(* IEC 61131-3 sources: JingjiangMoonbox/Application/Application/任务列表/Main_Task/GNS_MAP, 4 files *)

(* ---- KS_CreatGantryAxisInf.st ---- *)
(*@CES
Name=KS_CreatGantryAxisInf
Type=FunctionBlock
TypeGuid=6f9dac99-8de1-4efc-8465-68ac443b7d08
Guid=f41a9b20-4237-42b7-ab68-52a2ca659d0d
HasDeclaration=True
HasImplementation=True
*)
{DECLARATION}
FUNCTION KS_CreatGantryAxisInf : BOOL
(*获取龙门轴信息*)
VAR_INPUT
	(*输入*)
	i_pstStSysStationInf 	: POINTER TO StSysStationInf;
	(*输出*)
	i_pstStSysGantryAxisInf : POINTER TO StSysGantryAxisInf;
END_VAR
VAR
	in					: INT;
	pstStStationInf		: POINTER TO StStationInf;
	pstStGantryAxisInf	: POINTER TO StGantryAxisInf;
	(*龙门轴信息地址@索引为轴id,最大15*)
	(*每个轴2个龙门@二维数组里的1是版辊、2是网纹辊*)
	apstStGantryAxisInf	: ARRAY [1..20,1..2] OF POINTER TO StGantryAxisInf:=[40(0)];
	iGantryAxisNum		: INT := 0;(*龙门轴个数*)
	iMaxGantryAxisNum	: INT;
	iLogicAxisId		: INT;(*逻辑轴id*)
	iLogicAxisIdSuperPos: INT;(*叠加轴id*)
	iMoveType			: stEnumMoveType;(*运动类型*)
	iAxisId				: stEnumAxisId;
	iStaitonFuncId		: stEnumFuncId;
	iCoreId				: INT;
	iIndexTmp			: INT;(*数组索引*)
END_VAR
{IMPLEMENTATION}
IF i_pstStSysStationInf<>0 AND i_pstStSysGantryAxisInf<>0 THEN
	(*龙门组个数*)
	iMaxGantryAxisNum:=SIZEOF(i_pstStSysGantryAxisInf^.astGantryAxisInf)/SIZEOF(i_pstStSysGantryAxisInf^.astGantryAxisInf[1]);
	(*初始化*)
	FOR iN:=1 TO iMaxGantryAxisNum BY 1 DO
		KS_InitGantryAxisInf(ADR(i_pstStSysGantryAxisInf^.astGantryAxisInf[iN]));
	END_FOR
	(*从系统架构中找龙门轴*)
	FOR in:=1 TO i_pstStSysStationInf^.byStationNum BY 1 DO
		pstStStationInf:=ADR(i_pstStSysStationInf^.astStationInf[iN]);
		IF pstStStationInf^.xValid THEN
			iAxisId					:=pstStStationInf^.iAxisId;
			iLogicAxisId			:=pstStStationInf^.iLogicAxisId;
			iLogicAxisIdSuperPos	:=pstStStationInf^.iLogicAxisIdSuperPos;
			iMoveType				:=pstStStationInf^.iMoveType;
			iStaitonFuncId			:=pstStStationInf^.iFuncId;
			iCoreId					:=pstStStationInf^.iCoreId_LogicAxis;
			IF KS_IsUnitAxisId(iAxisId)THEN(*是色组*)
				IF iMoveType = MOVETYPE_GANTRY THEN(*龙门轴*)
					IF iStaitonFuncId = FUNCID_PRNROLLER_PRESSURE_M OR
						iStaitonFuncId = FUNCID_PRNROLLER_PRESSURE_G THEN(*印刷辊龙门*)
						iIndexTmp:=1;
					ELSE(*else都认为是网纹辊龙门*)
						iIndexTmp:=2;
					END_IF

					IF apstStGantryAxisInf[iAxisId,iIndexTmp] = 0 THEN
						iGantryAxisNum:=iGantryAxisNum+1;
						(*获取龙门轴需要的信息*)
						(*写入的结构体地址获取*)
						IF iGantryAxisNum<=iMaxGantryAxisNum THEN
							pstStGantryAxisInf:=ADR(i_pstStSysGantryAxisInf^.astGantryAxisInf[iGantryAxisNum]);
						ELSE(*超限了|退出*)
							EXIT;
						END_IF
						apstStGantryAxisInf[iAxisId,iIndexTmp]:=ADR(i_pstStSysGantryAxisInf^.astGantryAxisInf[iGantryAxisNum]);
					END_IF

					(*获取地址*)
					pstStGantryAxisInf:=apstStGantryAxisInf[iAxisId,iIndexTmp];
					IF pstStGantryAxisInf<>0 THEN(*地址合法*)
						pstStGantryAxisInf^.iAxisId:=iAxisId;
						pstStGantryAxisInf^.iCoreId:=iCoreId;(*龙门站必须是一个核|所以不用区分*)

						CASE iStaitonFuncId OF
							FUNCID_PRNROLLER_PRESSURE_M:(*版辊压力|操作侧@叠加轴id在m侧的数据里*)
								pstStGantryAxisInf^.iFuncId					:=FUNCID_PRNROLLER_GANTRY;
								pstStGantryAxisInf^.iLogicAxisId_M			:=iLogicAxisId;
								pstStGantryAxisInf^.iLogicAxisId_SuperPos	:=iLogicAxisIdSuperPos;
							FUNCID_PRNROLLER_PRESSURE_G:
								pstStGantryAxisInf^.iFuncId					:=FUNCID_PRNROLLER_GANTRY;
								pstStGantryAxisInf^.iLogicAxisId_G			:=pstStStationInf^.iLogicAxisId;
							FUNCID_NETROLLER_PRESSURE_M:(*网辊压力|操作侧@叠加轴id在m侧的数据里*)
								pstStGantryAxisInf^.iFuncId					:=FUNCID_NETROLLER_GANTRY;
								pstStGantryAxisInf^.iLogicAxisId_M			:=iLogicAxisId;
								pstStGantryAxisInf^.iLogicAxisId_SuperPos	:=iLogicAxisIdSuperPos;
							FUNCID_NETROLLER_PRESSURE_G:
								pstStGantryAxisInf^.iFuncId					:=FUNCID_NETROLLER_GANTRY;
								pstStGantryAxisInf^.iLogicAxisId_G			:=pstStStationInf^.iLogicAxisId;
						ELSE;(*不是压力的就不理会了*)
						END_CASE
					END_IF
				ELSE(*不是龙门轴不理会*);
				END_IF
			END_IF(*不是色组就不理会了*);
		END_IF
	END_FOR
	i_pstStSysGantryAxisInf^.byGantryAxisNum:=INT_TO_BYTE(iGantryAxisNum);

	(*非法值检测*)
	FOR iN:=1 TO iGantryAxisNum BY 1 DO
		pstStGantryAxisInf:=ADR(i_pstStSysGantryAxisInf^.astGantryAxisInf[iN]);
		pstStGantryAxisInf^.xValid:=TRUE;
		IF pstStGantryAxisInf^.iAxisId=-1 OR
			pstStGantryAxisInf^.iCoreId=-1 OR
			pstStGantryAxisInf^.iFuncId=FUNCID_NULL OR
			pstStGantryAxisInf^.iLogicAxisId_G=-1 OR
			pstStGantryAxisInf^.iLogicAxisId_M=-1 OR
			pstStGantryAxisInf^.iLogicAxisId_SuperPos=-1 THEN
			pstStGantryAxisInf^.xValid:=FALSE;
		END_IF
	END_FOR
END_IF

(* ---- KS_CreatMap.st ---- *)
(*@CES
Name=KS_CreatMap
Type=FunctionBlock
TypeGuid=6f9dac99-8de1-4efc-8465-68ac443b7d08
Guid=61e29dc5-e287-4a1a-b094-66cbd5c76957
HasDeclaration=True
HasImplementation=True
*)
{DECLARATION}
FUNCTION KS_CreatMap : BOOL
(*创建映射表@触发执行|初始化获取到了站列表后执行一次就行*)
(*对应关系参考站号定义、xml分配文件*)
(*新的架构需要同步修改KS_CreatStationIdMap\KS_GetLogicAxisInfByStationIdForMap*)
(*2026.5.20.140844 by liu.yt 调整接口为系统列表结构体*)
VAR_INPUT
	i_xEn					: BOOL;(*创建使能@事件触发*)
	i_xUseRealStation		: BOOL;(*使用实际站创建*)
	(*根据系统架构创建*)
	i_iMachineryType		: stEuumMachineryType;(*机器类型*)
(*
	i_xIsDualUwRw			: BOOL;(*双收双放机型|*)
	i_xIfOfIsGlink			: BOOL;(*收放牵是glink站*)
	i_xUwRwIsGlink			: BOOL;(*收放料是glink站*)
	i_xPrnPressureIsGlink	: BOOL;(*印刷辊的压力辊是glink站*)
	i_xNetPressureIsGlink	: BOOL;(*网纹辊的压力辊是glink站*)
*)

	(*系统中实际站信息*)
	i_byStationIdNum		: BYTE;(*站的个数*)
	//i_piStationIdList		: POINTER TO INT;(*站id列表*)
	i_pstStStationInfo_KS	: POINTER TO StStationInfo_KS;(*固高函数获取的系统站信息@2026.5.20.140838 by liu.yt*)
	(*输出列表*)
	i_pstStSysStationInf	: POINTER TO StSysStationInf;
END_VAR
VAR
	iN					: INT;
	iAxisId				: stEnumAxisId;
	piTmp				: POINTER TO INT;
	pwTmp				: POINTER TO WORD;
	iStationInflenth	: INT;
	iStationNum			: INT;(*站的个数*)
	iValidStationNum	: INT;(*有效站个数*)
	aiStationidList		: ARRAY [1..256] OF INT;
	wStationType		: WORD;(*站的类型*)
	awStationType		: ARRAY [1..256] OF WORD;(*2026.5.20.141316 by liu.yt*)
	pstStationInf		: POINTER TO StStationInf;
	iFuncId				: stEnumFuncId;(*只针对色组轴*)
	iMoveType			: stEnumMoveType;(*运动的类型也可以获取*)
	iStationId			: INT;
	iCoreId				: INT:=-1;
	iLogicAxisIdSuperPos: INT:=-1;
	iLogicAxisId		: INT:=-1;
	(*不同的机型必须要显式赋值*)
	(*色组数@默认写的是机组式柔印+4压力电机*)
	iUnitNum			: INT:=10;
	iMachineryType		: stEuumMachineryType;
END_VAR
{IMPLEMENTATION}
IF i_xEn THEN
	iStationInflenth:=SIZEOF(i_pstStSysStationInf^.astStationInf) /
						SIZEOF(i_pstStSysStationInf^.astStationInf[1]);
	iMachineryType:=i_iMachineryType;
	(*获取站列表和个数*)
	IF i_xUseRealStation THEN
		(*2026.5.20.141002 by liu.yt*)
		//iStationNum:=BYTE_TO_INT(i_byStationIdNum);
		(*piTmp:=i_piStationIdList;*)
		iStationNum:=i_pstStStationInfo_KS^.iStationNum;
		piTmp:=ADR(i_pstStStationInfo_KS^.aiStationId_List);
		pwTmp:=ADR(i_pstStStationInfo_KS^.awStation_Type);
		FOR iN:=1 TO iStationNum BY 1 DO
			(*列表获取@2026.5.20.141347 by liu.yt*)
			aiStationidList[iN]:=piTmp^;
			piTmp:=piTmp+SIZEOF(piTmp^);
			(*站类型获取@2026.5.20.141359 by liu.yt*)
			awStationType[iN]:=pwTmp^;
			pwTmp:=pwTmp+SIZEOF(pwTmp^);
		END_FOR
	ELSE
		iStationNum:=255(*iStationInflenth*);
		IF iStationNum<=255 THEN
			FOR iN:=1 TO iStationNum BY 1 DO
				aiStationidList[iN]:=iN;
			END_FOR
		END_IF
	END_IF
	(*初始化@结构体数据*)
	i_pstStSysStationInf^.byStationNum:=0;
	FOR iN:=1 TO iStationInflenth BY 1 DO
		pstStationInf:=ADR(i_pstStSysStationInf^.astStationInf[iN]);
		KS_InitStationInf(pstStationInf);
	END_FOR

	iValidStationNum:=0;
(*	IF NOT i_xIsDualUwRw THEN(*常规机型*)*)
		(*按照*)
		CASE iMachineryType OF
			MACHINERYTYPE_ROTOGRAVE:(*凹印机*);
			MACHINERYTYPE_FELXO_INLINE,(*机组式柔印*)
			MACHINERYTYPE_FELXO_INLINE_ONEBOTOMROLLER:(*机组式柔印@单底辊*)
				(*按照10色，带龙门压力，横向配置@压力轴的个数限制了最大色组数只能为10个*)
				iUnitNum:=10;(*4电机压力限制最大只能10色*)
				(*处理map*)
				FOR iN:=1 TO iStationNum BY 1 DO
					iStationId:=aiStationidList[iN];
					wStationType:=awStationType[iN];
					(*获取轴信息*)
					iAxisId:=KS_GetAxisInfByStationIdForMap(iStationId,ADR(iFuncId),ADR(iMoveType));
					(*站号在表里,就输出有效标志*)
					IF iAxisId<>AXISID_INVALID THEN
						IF iAxisId > iUnitNum AND iAxisId <= AXISID_15U THEN(*非法轴id就剔除*);
						ELSE;
							iValidStationNum:=iValidStationNum+1;
							IF iValidStationNum<=iStationInflenth THEN
								pstStationInf:=ADR(i_pstStSysStationInf^.astStationInf[iValidStationNum]);
								pstStationInf^.xValid:=TRUE;
								pstStationInf^.iAxisId:=iAxisId;
								pstStationInf^.iStationId:=iStationId;
								pstStationInf^.iFuncId:=iFuncId;
								pstStationInf^.iMoveType:=iMoveType;
								pstStationInf^.udiStationType:=WORD_TO_UDINT(wStationType);(*2026.5.20.161045 by liu.yt*)
								(*运控信息获取*)
								iLogicAxisId:=
									KS_GetLogicAxisInfByStationIdForMap(
												iStationId(*i_iStationId*),
												iMachineryType(*i_iMachineryType*),
												ADR(iCoreId)(*i_piCoreId*),
												ADR(iLogicAxisIdSuperPos)(*i_piLogicAxisIdSuperPos*));

								pstStationInf^.iCoreId_LogicAxis			:=iCoreId;
								pstStationInf^.iCoreId_LogicAxisSuperPos	:=iCoreId;
								pstStationInf^.iLogicAxisId					:=iLogicAxisId;
								pstStationInf^.iLogicAxisIdSuperPos			:=iLogicAxisIdSuperPos;
							ELSE;(*超过最大索引了*)
								iValidStationNum:=iStationInflenth;(*站个数最大就是数组长度*)
							END_IF
						END_IF
					END_IF
				END_FOR

			MACHINERYTYPE_FELXO_CL:(*卫星式柔印*);
			MACHINERYTYPE_OFFSET:(*胶印机*);
		ELSE;
		END_CASE
(*
	ELSE;
	END_IF
*)
	i_pstStSysStationInf^.byStationNum:=INT_TO_BYTE(iValidStationNum);
END_IF

//2025.12.27.142131 | + 机器类型搞个变量单独弄出来
g_iMachineryType := i_iMachineryType;

(* ---- KS_GetAxisIdForMotByStation_Gantry.st ---- *)
(*@CES
Name=KS_GetAxisIdForMotByStation_Gantry
Type=FunctionBlock
TypeGuid=6f9dac99-8de1-4efc-8465-68ac443b7d08
Guid=cde7d95e-737e-4f32-881d-821472d364d1
HasDeclaration=True
HasImplementation=True
*)
{DECLARATION}
FUNCTION KS_GetAxisIdForMotByStation_Gantry : BOOL
(*转换为火眼原来设计的数据项，并输出。方便程序移植*)
VAR_INPUT
	i_iStationId			: INT;
	i_piAxisId				: POINTER TO INT;(*逻辑轴id*)
	i_piTypeId				: POINTER TO ENUM_AXISTYPE;(*类型id*)
	i_piUnitId				: POINTER TO INT;(*色组id*)
	i_piCoreId				: POINTER TO INT;(*核id*)
	i_piGroupId			 	: POINTER TO INT;(*组id*)
	i_piAdjAxisId			: POINTER TO INT;(*调整轴id*)
	(*系统列表*)
	i_pstStSysStationInf	: POINTER TO StSysStationInf;
	i_pstStSysGantryAxisInf	: POINTER TO StSysGantryAxisInf;
END_VAR
VAR
	iN					:  INT;
	xResult				:  BOOL:=FALSE;
	iAxisId				:  INT:=-1;(*逻辑轴id*)
	iTypeId				:  ENUM_AXISTYPE:=TYPE_NULL;(*类型id*)
	iUnitId				:  INT:=-1;(*色组id*)
	iCoreId				:  INT:=-1;(*核id*)
	iGroupId			:  INT:=-1;(*组id*)
	iAdjAxisId			:  INT:=-1;(*调整轴id*)
	pstStStationInf 	:  POINTER TO StStationInf;
	pstStGantryAxisInf	:  POINTER TO StGantryAxisInf;
END_VAR

{IMPLEMENTATION}
IF i_pstStSysStationInf <>0 AND i_pstStSysGantryAxisInf <> 0 THEN
	IF i_iStationId>0 AND i_iStationId<255 THEN(*站号合法性判断*)
		FOR iN:=1 TO i_pstStSysStationInf^.byStationNum BY 1 DO
			pstStStationInf:=ADR(i_pstStSysStationInf^.astStationInf[iN]);
			IF pstStStationInf^.xValid THEN
				IF i_iStationId = pstStStationInf^.iStationId THEN(*找到了*)
					xResult:=TRUE;
					iAxisId:=pstStStationInf^.iLogicAxisId;(*逻辑轴id*)
					IF KS_IsUnitAxisId(pstStStationInf^.iAxisId) THEN(*检查是不是色组的枚举*)
						iUnitId:=pstStStationInf^.iAxisId;
					END_IF
					iCoreId:=pstStStationInf^.iCoreId_LogicAxis;(*核id*)
					iAdjAxisId:=pstStStationInf^.iLogicAxisIdSuperPos;(*叠加轴id*)
					EXIT;
				END_IF
			END_IF
		END_FOR
	END_IF

	(*type处理*)
	iTypeId:=TYPE_NULL;
	IF xResult THEN
		CASE pstStStationInf^.iAxisId OF
			AXISID_UWA:		iTypeId:=TYPE_UNWIND_A_I;
			AXISID_UWB:		iTypeId:=TYPE_UNWIND_B_I;
			AXISID_RWA:		iTypeId:=TYPE_REWIND_A_I;
			AXISID_RWB:		iTypeId:=TYPE_REWIND_B_I;
			AXISID_IF:		iTypeId:=TYPE_INFEED_I;
			AXISID_OF:		iTypeId:=TYPE_OUTFEED_I;
			AXISID_UWA_II:	iTypeId:=TYPE_UNWIND_A_II;
			AXISID_UWB_II:	iTypeId:=TYPE_UNWIND_B_II;
			AXISID_RWA_II:	iTypeId:=TYPE_REWIND_A_II;
			AXISID_RWB_II:	iTypeId:=TYPE_REWIND_B_II;
			AXISID_IF_II:	iTypeId:=TYPE_INFEED_II;
			AXISID_OF_II:	iTypeId:=TYPE_OUTFEED_II;
			AXISID_CENTER:  iTypeId:=TYPE_CENTRAL_I;(*只处理单系中心辊*)
		ELSE
			(*色组*)
			IF  KS_IsUnitAxisId(pstStStationInf^.iAxisId) THEN
				CASE pstStStationInf^.iFuncId OF
					FUNCID_PRNROLLER: 				iTypeId:=TYPE_UNIT_PRN;
					FUNCID_NETROLLER: 				iTypeId:=TYPE_UNIT_NET;
					FUNCID_BOTTOMROLLER: 			iTypeId:=TYPE_UNIT_BOTTOM;
					FUNCID_PRNROLLER_PRESSURE_M: 	iTypeId:=TYPE_UNIT_PRN_PRESS_MASTER;
					FUNCID_PRNROLLER_PRESSURE_G: 	iTypeId:=TYPE_UNIT_PRN_PRESS_G;
					FUNCID_NETROLLER_PRESSURE_M: 	iTypeId:=TYPE_UNIT_NET_PRESS_MASTER;
					FUNCID_NETROLLER_PRESSURE_G: 	iTypeId:=TYPE_UNIT_NET_PRESS_G;
					FUNCID_HORZ: 					iTypeId:=TYPE_UNIT_HORIZ;
				ELSE;
				END_CASE
			END_IF
		END_CASE
	END_IF

	//龙门处理
	FOR iN:=1 TO i_pstStSysGantryAxisInf^.byGantryAxisNum BY 1 DO
		pstStGantryAxisInf := ADR(i_pstStSysGantryAxisInf^.astGantryAxisInf[iN]);
		IF  pstStGantryAxisInf^.xValid THEN
			IF iUnitId = pstStGantryAxisInf^.iAxisId THEN
				IF pstStGantryAxisInf^.iFuncId = FUNCID_PRNROLLER_GANTRY THEN
					IF iTypeId = TYPE_UNIT_PRN_PRESS_MASTER OR iTypeId = TYPE_UNIT_PRN_PRESS_G THEN
						iGroupId := iN;
						EXIT;
					END_IF
				ELSIF pstStGantryAxisInf^.iFuncId = FUNCID_NETROLLER_GANTRY THEN
					IF iTypeId = TYPE_UNIT_NET_PRESS_MASTER OR iTypeId = TYPE_UNIT_NET_PRESS_G THEN
						iGroupId := iN;
						EXIT;
					END_IF
				END_IF
			END_IF
		END_IF
	END_FOR
END_IF

IF i_piAxisId<>0 THEN
	i_piAxisId^:=iAxisId;
END_IF
IF i_piTypeId<>0 THEN
	i_piTypeId^:=iTypeId;
END_IF
IF i_piUnitId<>0 THEN
	i_piUnitId^:=iUnitId;
END_IF
IF i_piCoreId<>0 THEN
	i_piCoreId^:=iCoreId;
END_IF
IF i_piGroupId<>0 THEN
	i_piGroupId^:=iGroupId;
END_IF
IF i_piAdjAxisId<>0 THEN
	i_piAdjAxisId^:=iAdjAxisId;
END_IF
KS_GetAxisIdForMotByStation_Gantry:=xResult;

(* ---- KS_GetAxisIdForMotByStation_V2.st ---- *)
(*@CES
Name=KS_GetAxisIdForMotByStation_V2
Type=FunctionBlock
TypeGuid=6f9dac99-8de1-4efc-8465-68ac443b7d08
Guid=c5880d4f-2cd9-4162-8439-8609b06a0444
HasDeclaration=True
HasImplementation=True
*)
{DECLARATION}
FUNCTION KS_GetAxisIdForMotByStation_V2 : BOOL
(*转换为火眼原来设计的数据项，并输出。方便程序移植*)
VAR_INPUT
	i_iStationId			: INT;
	i_piAxisId				: POINTER TO INT;(*逻辑轴id*)
	i_piTypeId				: POINTER TO ENUM_AXISTYPE;(*类型id*)
	i_piUnitId				: POINTER TO INT;(*色组id*)
	i_piCoreId				: POINTER TO INT;(*核id*)
	i_piGroupId			 	: POINTER TO INT;(*组id*)
	i_piAdjAxisId			: POINTER TO INT;(*调整轴id*)
	(*系统列表*)
	i_pstStSysStationInf	: POINTER TO StSysStationInf;
END_VAR
VAR
	iN					:  INT;
	xResult				:  BOOL:=FALSE;
	iAxisId				:  INT:=-1;(*逻辑轴id*)
	iTypeId				:  ENUM_AXISTYPE:=TYPE_NULL;(*类型id*)
	iUnitId				:  INT:=-1;(*色组id*)
	iCoreId				:  INT:=-1;(*核id*)
	iGroupId			:  INT:=-1;(*组id*)
	iAdjAxisId			:  INT:=-1;(*调整轴id*)
	pstStStationInf		:  POINTER TO StStationInf;
END_VAR
{IMPLEMENTATION}
IF i_pstStSysStationInf <>0 THEN
	IF i_iStationId>0 AND i_iStationId<255 THEN(*站号合法性判断*)
		FOR iN:=1 TO i_pstStSysStationInf^.byStationNum BY 1 DO
			pstStStationInf:=ADR(i_pstStSysStationInf^.astStationInf[iN]);
			IF pstStStationInf^.xValid THEN
				IF i_iStationId = pstStStationInf^.iStationId THEN(*找到了*)
					xResult:=TRUE;
					iAxisId:=pstStStationInf^.iLogicAxisId;(*逻辑轴id*)
					IF KS_IsUnitAxisId(pstStStationInf^.iAxisId) THEN(*检查是不是色组的枚举*)
						iUnitId:=pstStStationInf^.iAxisId;
					END_IF
					iCoreId:=pstStStationInf^.iCoreId_LogicAxis;(*核id*)
					iAdjAxisId:=pstStStationInf^.iLogicAxisIdSuperPos;(*叠加轴id*)
					EXIT;
				END_IF
			END_IF
		END_FOR
	END_IF

	(*type处理*)
	iTypeId:=TYPE_NULL;
	IF xResult THEN
		CASE pstStStationInf^.iAxisId OF
			AXISID_UWA:		iTypeId:=TYPE_UNWIND_A_I;
			AXISID_UWB:		iTypeId:=TYPE_UNWIND_B_I;
			AXISID_RWA:		iTypeId:=TYPE_REWIND_A_I;
			AXISID_RWB:		iTypeId:=TYPE_REWIND_B_I;
			AXISID_IF:		iTypeId:=TYPE_INFEED_I;
			AXISID_OF:		iTypeId:=TYPE_OUTFEED_I;
			AXISID_UWA_II:	iTypeId:=TYPE_UNWIND_A_II;
			AXISID_UWB_II:	iTypeId:=TYPE_UNWIND_B_II;
			AXISID_RWA_II:	iTypeId:=TYPE_REWIND_A_II;
			AXISID_RWB_II:	iTypeId:=TYPE_REWIND_B_II;
			AXISID_IF_II:	iTypeId:=TYPE_INFEED_II;
			AXISID_OF_II:	iTypeId:=TYPE_OUTFEED_II;
			AXISID_CENTER:  iTypeId:=TYPE_CENTRAL_I;(*只处理单系中心辊*)
		ELSE
			(*色组*)
			IF  KS_IsUnitAxisId(pstStStationInf^.iAxisId) THEN
				CASE pstStStationInf^.iFuncId OF
					FUNCID_CONTROL:					iTypeId:=TYPE_UNIT_CTL;(*2026.5.20.135932 by liu.yt*)
					FUNCID_PRNROLLER: 				iTypeId:=TYPE_UNIT_PRN;
					FUNCID_NETROLLER: 				iTypeId:=TYPE_UNIT_NET;
					FUNCID_BOTTOMROLLER: 			iTypeId:=TYPE_UNIT_BOTTOM;
					FUNCID_PRNROLLER_PRESSURE_M: 	iTypeId:=TYPE_UNIT_PRN_PRESS_MASTER;
					FUNCID_PRNROLLER_PRESSURE_G: 	iTypeId:=TYPE_UNIT_PRN_PRESS_G;
					FUNCID_NETROLLER_PRESSURE_M: 	iTypeId:=TYPE_UNIT_NET_PRESS_MASTER;
					FUNCID_NETROLLER_PRESSURE_G: 	iTypeId:=TYPE_UNIT_NET_PRESS_G;
					FUNCID_HORZ: 					iTypeId:=TYPE_UNIT_HORIZ;
				ELSE;
				END_CASE
			END_IF
		END_CASE
	END_IF
END_IF

IF i_piAxisId<>0 THEN
	i_piAxisId^:=iAxisId;
END_IF
IF i_piTypeId<>0 THEN
	i_piTypeId^:=iTypeId;
END_IF
IF i_piUnitId<>0 THEN
	i_piUnitId^:=iUnitId;
END_IF
IF i_piCoreId<>0 THEN
	i_piCoreId^:=iCoreId;
END_IF
IF i_piGroupId<>0 THEN
	i_piGroupId^:=iGroupId;
END_IF
IF i_piAdjAxisId<>0 THEN
	i_piAdjAxisId^:=iAdjAxisId;
END_IF
KS_GetAxisIdForMotByStation_V2:=xResult;
